(* IEC 61131-3 sources: plcassist-cli/packages/volt-lsp-iec/test-corpus/awa-palletizer/Device/Plc Logic/Application/Library Manager/SysFile, 21 files *)

(* ---- SYSFILECLOSE.fun ---- *)
FUNCTION SYSFILECLOSE : RTS_IEC_RESULT
VAR_INPUT
	HFILE : RTS_IEC_HANDLE;
END_VAR
END_FUNCTION

(* ---- SYSFILECOPY.fun ---- *)
FUNCTION SYSFILECOPY : RTS_IEC_RESULT
VAR_INPUT
	SZDESTFILENAME : REFERENCE TO STRING;
	SZSOURCEFILENAME : REFERENCE TO STRING;
	PULCOPIED : POINTER TO __XWORD;
END_VAR
END_FUNCTION

(* ---- SYSFILEDELETE.fun ---- *)
FUNCTION SYSFILEDELETE : RTS_IEC_RESULT
VAR_INPUT
	SZFILENAME : REFERENCE TO STRING;
END_VAR
END_FUNCTION

(* ---- SYSFILEDELETEBYHANDLE.fun ---- *)
FUNCTION SYSFILEDELETEBYHANDLE : RTS_IEC_RESULT
VAR_INPUT
	HFILE : RTS_IEC_HANDLE;
END_VAR
END_FUNCTION

(* ---- SYSFILEEOF.fun ---- *)
FUNCTION SYSFILEEOF : RTS_IEC_RESULT
VAR_INPUT
	HFILE : RTS_IEC_HANDLE;
END_VAR
END_FUNCTION

(* ---- SYSFILEFLUSH.fun ---- *)
FUNCTION SYSFILEFLUSH : RTS_IEC_RESULT
VAR_INPUT
	HFILE : RTS_IEC_HANDLE;
END_VAR
END_FUNCTION

(* ---- SYSFILEGETNAME.fun ---- *)
FUNCTION SYSFILEGETNAME : POINTER TO STRING
VAR_INPUT
	HFILE : RTS_IEC_HANDLE;
END_VAR
END_FUNCTION

(* ---- SYSFILEGETNAME2.fun ---- *)
FUNCTION SYSFILEGETNAME2 : POINTER TO STRING
VAR_INPUT
	HFILE : RTS_IEC_HANDLE;
	PRESULT : POINTER TO RTS_IEC_RESULT;
END_VAR
END_FUNCTION

(* ---- SYSFILEGETPATH.fun ---- *)
FUNCTION SYSFILEGETPATH : RTS_IEC_RESULT
VAR_INPUT
	SZFILENAME : REFERENCE TO STRING;
	DIMAXLEN : DINT;
END_VAR
VAR_IN_OUT
	SZPATH : STRING;
END_VAR
END_FUNCTION

(* ---- SYSFILEGETPOS.fun ---- *)
FUNCTION SYSFILEGETPOS : RTS_IEC_RESULT
VAR_INPUT
	HFILE : RTS_IEC_HANDLE;
	PULPOS : POINTER TO __XWORD;
END_VAR
END_FUNCTION

(* ---- SYSFILEGETSIZE.fun ---- *)
FUNCTION SYSFILEGETSIZE : __XWORD
VAR_INPUT
	SZFILENAME : REFERENCE TO STRING;
	PRESULT : POINTER TO RTS_IEC_RESULT;
END_VAR
END_FUNCTION

(* ---- SYSFILEGETSIZEBYHANDLE.fun ---- *)
FUNCTION SYSFILEGETSIZEBYHANDLE : __XWORD
VAR_INPUT
	HFILE : RTS_IEC_HANDLE;
	PRESULT : POINTER TO RTS_IEC_RESULT;
END_VAR
END_FUNCTION

(* ---- SYSFILEGETSTATUS.fun ---- *)
FUNCTION SYSFILEGETSTATUS : SYS_FILE_STATUS
VAR_INPUT
	HFILE : RTS_IEC_HANDLE;
END_VAR
END_FUNCTION

(* ---- SYSFILEGETSTATUS2.fun ---- *)
FUNCTION SYSFILEGETSTATUS2 : SYS_FILE_STATUS
VAR_INPUT
	HFILE : RTS_IEC_HANDLE;
	PRESULT : POINTER TO RTS_IEC_RESULT;
END_VAR
END_FUNCTION

(* ---- SYSFILEGETTIME.fun ---- *)
FUNCTION SYSFILEGETTIME : RTS_IEC_RESULT
VAR_INPUT
	SZFILENAME : REFERENCE TO STRING;
	PTFILETIME : POINTER TO SYS_FILETIME;
END_VAR
END_FUNCTION

(* ---- SYSFILEOPEN.fun ---- *)
FUNCTION SYSFILEOPEN : RTS_IEC_HANDLE
VAR_INPUT
	SZFILE : REFERENCE TO STRING;
	AM : ACCESS_MODE;
	PRESULT : POINTER TO RTS_IEC_RESULT;
END_VAR
END_FUNCTION

(* ---- SYSFILEREAD.fun ---- *)
FUNCTION SYSFILEREAD : __XWORD
VAR_INPUT
	HFILE : RTS_IEC_HANDLE;
	PBYBUFFER : POINTER TO BYTE;
	ULSIZE : __XWORD;
	PRESULT : POINTER TO RTS_IEC_RESULT;
END_VAR
END_FUNCTION

(* ---- SYSFILERENAME.fun ---- *)
FUNCTION SYSFILERENAME : RTS_IEC_RESULT
VAR_INPUT
	SZOLDFILENAME : REFERENCE TO STRING;
	SZNEWFILENAME : REFERENCE TO STRING;
END_VAR
END_FUNCTION

(* ---- SYSFILESETPOS.fun ---- *)
FUNCTION SYSFILESETPOS : RTS_IEC_RESULT
VAR_INPUT
	HFILE : RTS_IEC_HANDLE;
	ULOFFSET : __XWORD;
END_VAR
END_FUNCTION

(* ---- SYSFILETRUNCATE.fun ---- *)
FUNCTION SYSFILETRUNCATE : RTS_IEC_RESULT
VAR_INPUT
	HFILE : RTS_IEC_HANDLE;
	ULSIZENEW : __XWORD;
END_VAR
END_FUNCTION

(* ---- SYSFILEWRITE.fun ---- *)
FUNCTION SYSFILEWRITE : __XWORD
VAR_INPUT
	HFILE : RTS_IEC_HANDLE;
	PBYBUFFER : POINTER TO BYTE;
	ULSIZE : __XWORD;
	PRESULT : POINTER TO RTS_IEC_RESULT;
END_VAR
END_FUNCTION
